(* IEC 61131-3 sources: plc-st-coding-agent/progress/evidence/f14_v11_public_20261113/jobs/custom_minimax-m27, 8 files *)

(* ---- public-easy-01.candidate_01.st ---- *)
(* ENGINEERING_CONTRACT
+--------------------------------------------------------------------------------------+
| Output             | Activation                | Retention | Reset/Deactivation    | Units |
|--------------------|---------------------------|-----------|-----------------------|-------|
| Pump_Motor         | bottleSensor in IDLE      | Hold      | cleaningConfirmButton | BOOL  |
| Filling_Valve      | cleaningConfirmButton     | Hold      | fillingConfirmButton  | BOOL  |
| Capping_Machine    | fillingConfirmButton      | Hold      | cappingConfirmButton  | BOOL  |
| Packing_Machine    | cappingConfirmButton      | Hold      | packingConfirmButton  | BOOL  |
| Completion_Light   | packingConfirmButton      | Hold      | finishedButton        | BOOL  |
+--------------------------------------------------------------------------------------+
| State Machine: IDLE->CLEANING->FILLING->CAPPING->PACKING->COMPLETED->IDLE           |
| All confirm inputs use R_TRIG for edge detection (same-scan priority preserved).     |
| Outputs are combinational to their active state; no edge memory needed.              |
| finishedButton only resets from COMPLETED state (PUB008).                            |
+--------------------------------------------------------------------------------------+
*)
(* CONTRACT_RULES [{"kind":"hold_until_reset","output":"Completion_Light","set_input":"packingConfirmButton","reset_input":"finishedButton"}] *)
FUNCTION_BLOCK BottleFillingLine
VAR_INPUT
    bottleSensor          : BOOL;
    cleaningConfirmButton : BOOL;
    fillingConfirmButton  : BOOL;
    cappingConfirmButton  : BOOL;
    packingConfirmButton  : BOOL;
    finishedButton        : BOOL;
END_VAR
VAR_OUTPUT
    Pump_Motor      : BOOL;
    Filling_Valve   : BOOL;
    Capping_Machine : BOOL;
    Packing_Machine : BOOL;
    Completion_Light: BOOL;
END_VAR
VAR
    eState : INT;
    IDLE      : INT := 0;
    CLEANING  : INT := 1;
    FILLING   : INT := 2;
    CAPPING   : INT := 3;
    PACKING   : INT := 4;
    COMPLETED : INT := 5;

    trigBottle   : R_TRIG;
    trigClean    : R_TRIG;
    trigFill     : R_TRIG;
    trigCap      : R_TRIG;
    trigPack     : R_TRIG;
    trigFinished : R_TRIG;
END_VAR

// Detect rising edges for all button inputs
trigBottle(CLK := bottleSensor);
trigClean(CLK := cleaningConfirmButton);
trigFill(CLK := fillingConfirmButton);
trigCap(CLK := cappingConfirmButton);
trigPack(CLK := packingConfirmButton);
trigFinished(CLK := finishedButton);

// State machine transitions
CASE eState OF
    IDLE:
        IF trigBottle.Q THEN
            eState := CLEANING;
        END_IF;

    CLEANING:
        IF trigClean.Q THEN
            eState := FILLING;
        END_IF;

    FILLING:
        IF trigFill.Q THEN
            eState := CAPPING;
        END_IF;

    CAPPING:
        IF trigCap.Q THEN
            eState := PACKING;
        END_IF;

    PACKING:
        IF trigPack.Q THEN
            eState := COMPLETED;
        END_IF;

    COMPLETED:
        IF trigFinished.Q THEN
            eState := IDLE;
        END_IF;
END_CASE;

// Output control based on current state
Pump_Motor       := (eState = CLEANING);
Filling_Valve    := (eState = FILLING);
Capping_Machine  := (eState = CAPPING);
Packing_Machine  := (eState = PACKING);
Completion_Light := (eState = COMPLETED);

END_FUNCTION_BLOCK

(* ---- public-easy-01.candidate_02.st ---- *)
(* ENGINEERING_CONTRACT
+--------------------------------------------------------------------------------------+
| Output             | Activation                | Retention | Reset/Deactivation    | Units |
|--------------------|---------------------------|-----------|-----------------------|-------|
| Pump_Motor         | bottleSensor in IDLE      | Hold      | cleaningConfirmButton | BOOL  |
| Filling_Valve      | cleaningConfirmButton     | Hold      | fillingConfirmButton  | BOOL  |
| Capping_Machine    | fillingConfirmButton      | Hold      | cappingConfirmButton  | BOOL  |
| Packing_Machine    | cappingConfirmButton      | Hold      | packingConfirmButton  | BOOL  |
| Completion_Light   | packingConfirmButton      | Hold      | finishedButton        | BOOL  |
+--------------------------------------------------------------------------------------+
| State Machine: IDLE->CLEANING->FILLING->CAPPING->PACKING->COMPLETED->IDLE           |
| All confirm inputs use R_TRIG for edge detection (same-scan priority preserved).     |
| Outputs are combinational to their active state; no edge memory needed.              |
| finishedButton only resets from COMPLETED state (PUB008).                            |
+--------------------------------------------------------------------------------------+
*)
(* CONTRACT_RULES [{"kind":"hold_until_reset","output":"Completion_Light","set_input":"packingConfirmButton","reset_input":"finishedButton"}] *)
FUNCTION_BLOCK BottleFillingLine
VAR_INPUT
    bottleSensor          : BOOL;
    cleaningConfirmButton : BOOL;
    fillingConfirmButton  : BOOL;
    cappingConfirmButton  : BOOL;
    packingConfirmButton  : BOOL;
    finishedButton        : BOOL;
END_VAR
VAR_OUTPUT
    Pump_Motor      : BOOL;
    Filling_Valve   : BOOL;
    Capping_Machine : BOOL;
    Packing_Machine : BOOL;
    Completion_Light: BOOL;
END_VAR
VAR
    eState : INT;

    trigBottle   : R_TRIG;
    trigClean    : R_TRIG;
    trigFill     : R_TRIG;
    trigCap      : R_TRIG;
    trigPack     : R_TRIG;
    trigFinished : R_TRIG;
END_VAR
VAR CONSTANT
    IDLE      : INT := 0;
    CLEANING  : INT := 1;
    FILLING   : INT := 2;
    CAPPING   : INT := 3;
    PACKING   : INT := 4;
    COMPLETED : INT := 5;
END_VAR

// Detect rising edges for all button inputs
trigBottle(CLK := bottleSensor);
trigClean(CLK := cleaningConfirmButton);
trigFill(CLK := fillingConfirmButton);
trigCap(CLK := cappingConfirmButton);
trigPack(CLK := packingConfirmButton);
trigFinished(CLK := finishedButton);

// State machine transitions
CASE eState OF
    IDLE:
        IF trigBottle.Q THEN
            eState := CLEANING;
        END_IF;

    CLEANING:
        IF trigClean.Q THEN
            eState := FILLING;
        END_IF;

    FILLING:
        IF trigFill.Q THEN
            eState := CAPPING;
        END_IF;

    CAPPING:
        IF trigCap.Q THEN
            eState := PACKING;
        END_IF;

    PACKING:
        IF trigPack.Q THEN
            eState := COMPLETED;
        END_IF;

    COMPLETED:
        IF trigFinished.Q THEN
            eState := IDLE;
        END_IF;
END_CASE;

// Output control based on current state
Pump_Motor       := (eState = CLEANING);
Filling_Valve    := (eState = FILLING);
Capping_Machine  := (eState = CAPPING);
Packing_Machine  := (eState = PACKING);
Completion_Light := (eState = COMPLETED);

END_FUNCTION_BLOCK

(* ---- public-easy-01.raw_candidate_01.st ---- *)
(* ENGINEERING_CONTRACT
+--------------------------------------------------------------------------------------+
| Output             | Activation                | Retention | Reset/Deactivation    | Units |
|--------------------|---------------------------|-----------|-----------------------|-------|
| Pump_Motor         | bottleSensor in IDLE      | Hold      | cleaningConfirmButton | BOOL  |
| Filling_Valve      | cleaningConfirmButton     | Hold      | fillingConfirmButton  | BOOL  |
| Capping_Machine    | fillingConfirmButton      | Hold      | cappingConfirmButton  | BOOL  |
| Packing_Machine    | cappingConfirmButton      | Hold      | packingConfirmButton  | BOOL  |
| Completion_Light   | packingConfirmButton      | Hold      | finishedButton        | BOOL  |
+--------------------------------------------------------------------------------------+
| State Machine: IDLE->CLEANING->FILLING->CAPPING->PACKING->COMPLETED->IDLE           |
| All confirm inputs use R_TRIG for edge detection (same-scan priority preserved).     |
| Outputs are combinational to their active state; no edge memory needed.              |
| finishedButton only resets from COMPLETED state (PUB008).                            |
+--------------------------------------------------------------------------------------+
*)
(* CONTRACT_RULES [{"kind":"hold_until_reset","output":"Completion_Light","set_input":"packingConfirmButton","reset_input":"finishedButton"}] *)
FUNCTION_BLOCK BottleFillingLine
VAR_INPUT
    bottleSensor          : BOOL;
    cleaningConfirmButton : BOOL;
    fillingConfirmButton  : BOOL;
    cappingConfirmButton  : BOOL;
    packingConfirmButton  : BOOL;
    finishedButton        : BOOL;
END_VAR
VAR_OUTPUT
    Pump_Motor      : BOOL;
    Filling_Valve   : BOOL;
    Capping_Machine : BOOL;
    Packing_Machine : BOOL;
    Completion_Light: BOOL;
END_VAR
VAR
    eState : INT;
    IDLE      : INT := 0;
    CLEANING  : INT := 1;
    FILLING   : INT := 2;
    CAPPING   : INT := 3;
    PACKING   : INT := 4;
    COMPLETED : INT := 5;

    trigBottle   : R_TRIG;
    trigClean    : R_TRIG;
    trigFill     : R_TRIG;
    trigCap      : R_TRIG;
    trigPack     : R_TRIG;
    trigFinished : R_TRIG;
END_VAR

// Detect rising edges for all button inputs
trigBottle(CLK := bottleSensor);
trigClean(CLK := cleaningConfirmButton);
trigFill(CLK := fillingConfirmButton);
trigCap(CLK := cappingConfirmButton);
trigPack(CLK := packingConfirmButton);
trigFinished(CLK := finishedButton);

// State machine transitions
CASE eState OF
    IDLE:
        IF trigBottle.Q THEN
            eState := CLEANING;
        END_IF;

    CLEANING:
        IF trigClean.Q THEN
            eState := FILLING;
        END_IF;

    FILLING:
        IF trigFill.Q THEN
            eState := CAPPING;
        END_IF;

    CAPPING:
        IF trigCap.Q THEN
            eState := PACKING;
        END_IF;

    PACKING:
        IF trigPack.Q THEN
            eState := COMPLETED;
        END_IF;

    COMPLETED:
        IF trigFinished.Q THEN
            eState := IDLE;
        END_IF;
END_CASE;

// Output control based on current state
Pump_Motor       := (eState = CLEANING);
Filling_Valve    := (eState = FILLING);
Capping_Machine  := (eState = CAPPING);
Packing_Machine  := (eState = PACKING);
Completion_Light := (eState = COMPLETED);

END_FUNCTION_BLOCK

(* ---- public-easy-01.raw_candidate_02.st ---- *)
(* ENGINEERING_CONTRACT
+--------------------------------------------------------------------------------------+
| Output             | Activation                | Retention | Reset/Deactivation    | Units |
|--------------------|---------------------------|-----------|-----------------------|-------|
| Pump_Motor         | bottleSensor in IDLE      | Hold      | cleaningConfirmButton | BOOL  |
| Filling_Valve      | cleaningConfirmButton     | Hold      | fillingConfirmButton  | BOOL  |
| Capping_Machine    | fillingConfirmButton      | Hold      | cappingConfirmButton  | BOOL  |
| Packing_Machine    | cappingConfirmButton      | Hold      | packingConfirmButton  | BOOL  |
| Completion_Light   | packingConfirmButton      | Hold      | finishedButton        | BOOL  |
+--------------------------------------------------------------------------------------+
| State Machine: IDLE->CLEANING->FILLING->CAPPING->PACKING->COMPLETED->IDLE           |
| All confirm inputs use R_TRIG for edge detection (same-scan priority preserved).     |
| Outputs are combinational to their active state; no edge memory needed.              |
| finishedButton only resets from COMPLETED state (PUB008).                            |
+--------------------------------------------------------------------------------------+
*)
(* CONTRACT_RULES [{"kind":"hold_until_reset","output":"Completion_Light","set_input":"packingConfirmButton","reset_input":"finishedButton"}] *)
FUNCTION_BLOCK BottleFillingLine
VAR_INPUT
    bottleSensor          : BOOL;
    cleaningConfirmButton : BOOL;
    fillingConfirmButton  : BOOL;
    cappingConfirmButton  : BOOL;
    packingConfirmButton  : BOOL;
    finishedButton        : BOOL;
END_VAR
VAR_OUTPUT
    Pump_Motor      : BOOL;
    Filling_Valve   : BOOL;
    Capping_Machine : BOOL;
    Packing_Machine : BOOL;
    Completion_Light: BOOL;
END_VAR
VAR
    eState : INT;

    trigBottle   : R_TRIG;
    trigClean    : R_TRIG;
    trigFill     : R_TRIG;
    trigCap      : R_TRIG;
    trigPack     : R_TRIG;
    trigFinished : R_TRIG;
END_VAR
VAR CONSTANT
    IDLE      : INT := 0;
    CLEANING  : INT := 1;
    FILLING   : INT := 2;
    CAPPING   : INT := 3;
    PACKING   : INT := 4;
    COMPLETED : INT := 5;
END_VAR

// Detect rising edges for all button inputs
trigBottle(CLK := bottleSensor);
trigClean(CLK := cleaningConfirmButton);
trigFill(CLK := fillingConfirmButton);
trigCap(CLK := cappingConfirmButton);
trigPack(CLK := packingConfirmButton);
trigFinished(CLK := finishedButton);

// State machine transitions
CASE eState OF
    IDLE:
        IF trigBottle.Q THEN
            eState := CLEANING;
        END_IF;

    CLEANING:
        IF trigClean.Q THEN
            eState := FILLING;
        END_IF;

    FILLING:
        IF trigFill.Q THEN
            eState := CAPPING;
        END_IF;

    CAPPING:
        IF trigCap.Q THEN
            eState := PACKING;
        END_IF;

    PACKING:
        IF trigPack.Q THEN
            eState := COMPLETED;
        END_IF;

    COMPLETED:
        IF trigFinished.Q THEN
            eState := IDLE;
        END_IF;
END_CASE;

// Output control based on current state
Pump_Motor       := (eState = CLEANING);
Filling_Valve    := (eState = FILLING);
Capping_Machine  := (eState = CAPPING);
Packing_Machine  := (eState = PACKING);
Completion_Light := (eState = COMPLETED);

END_FUNCTION_BLOCK

(* ---- public-easy-02.candidate_01.st ---- *)
(* ENGINEERING_CONTRACT:
 * - Inputs: value (DWORD, 32-bit), sampled every scan cycle
 * - Rising edge: prev=0 AND current=1 → risingBits = value AND NOT prevValue
 * - Falling edge: prev=1 AND current=0 → fallingBits = NOT value AND prevValue
 * - hasChanged: retention until next scan, set when value <> prevValue
 * - hasRisingEdges: combinational, true when risingBits <> 0
 * - hasFallingEdges: combinational, true when fallingBits <> 0
 * - risingBits/fallingBits: stored per-bit edge indicators, latching across scans
 * - noOfRisingBits/noOfFallingBits: USINT count of set bits in edge bitmasks
 * - Units: bit positions 0-31, counts 0-32
 * - Initialization: prevValue defaults to 0; first scan treats 0→1 as rising edges
 * - No explicit reset; state evolves per scan with prevValue update
 * - PUB001: Input value, edge detection logic, output reporting
 *)

(* CONTRACT_RULES [] *)

FUNCTION_BLOCK FB_DualWordEdgeDetection
VAR_INPUT
    value : DWORD;
END_VAR

VAR_OUTPUT
    hasChanged      : BOOL;
    hasRisingEdges  : BOOL;
    risingBits      : DWORD;
    noOfRisingBits  : USINT;
    hasFallingEdges : BOOL;
    fallingBits     : DWORD;
    noOfFallingBits : USINT;
END_VAR

VAR
    prevValue : DWORD;
END_VAR

VAR_TEMP
    tmp_i     : USINT;
END_VAR

    // Detect rising edges: current=1 AND previous=0
    risingBits := value AND NOT prevValue;

    // Detect falling edges: previous=1 AND current=0
    fallingBits := NOT value AND prevValue;

    // Report change detection
    hasChanged := value <> prevValue;

    // Report edge occurrence flags
    hasRisingEdges := risingBits <> 0;
    hasFallingEdges := fallingBits <> 0;

    // Count rising bits (0-32)
    noOfRisingBits := 0;
    FOR tmp_i := 0 TO 31 DO
        IF (risingBits AND (1 SHL tmp_i)) <> 0 THEN
            noOfRisingBits := noOfRisingBits + 1;
        END_IF;
    END_FOR;

    // Count falling bits (0-32)
    noOfFallingBits := 0;
    FOR tmp_i := 0 TO 31 DO
        IF (fallingBits AND (1 SHL tmp_i)) <> 0 THEN
            noOfFallingBits := noOfFallingBits + 1;
        END_IF;
    END_FOR;

    // Store current value for next scan comparison
    prevValue := value;
END_FUNCTION_BLOCK

(* ---- public-easy-02.candidate_02.st ---- *)
(* ENGINEERING_CONTRACT:
 * - Inputs: value (DWORD, 32-bit), sampled every scan cycle
 * - Rising edge: prev=0 AND current=1 → risingBits = value AND NOT prevValue
 * - Falling edge: prev=1 AND current=0 → fallingBits = NOT value AND prevValue
 * - hasChanged: retention until next scan, set when value <> prevValue
 * - hasRisingEdges: combinational, true when risingBits <> 0
 * - hasFallingEdges: combinational, true when fallingBits <> 0
 * - risingBits/fallingBits: stored per-bit edge indicators, latching across scans
 * - noOfRisingBits/noOfFallingBits: USINT count of set bits in edge bitmasks
 * - Units: bit positions 0-31, counts 0-32
 * - Initialization: prevValue defaults to 0; first scan treats 0→1 as rising edges
 * - No explicit reset; state evolves per scan with prevValue update
 * - PUB001: Input value, edge detection logic, output reporting
 *)

(* CONTRACT_RULES [] *)

FUNCTION_BLOCK FB_DualWordEdgeDetection
VAR_INPUT
    value : DWORD;
END_VAR

VAR_OUTPUT
    hasChanged      : BOOL;
    hasRisingEdges  : BOOL;
    risingBits      : DWORD;
    noOfRisingBits  : USINT;
    hasFallingEdges : BOOL;
    fallingBits     : DWORD;
    noOfFallingBits : USINT;
END_VAR

VAR
    prevValue : DWORD;
END_VAR

VAR_TEMP
    tmp_i     : USINT;
END_VAR

    // Detect rising edges: current=1 AND previous=0
    risingBits := value AND NOT prevValue;

    // Detect falling edges: previous=1 AND current=0
    fallingBits := NOT value AND prevValue;

    // Report change detection
    hasChanged := value <> prevValue;

    // Report edge occurrence flags
    hasRisingEdges := risingBits <> 0;
    hasFallingEdges := fallingBits <> 0;

    // Count rising bits (0-32)
    noOfRisingBits := 0;
    FOR tmp_i := 0 TO 31 DO
        IF (risingBits AND SHL(1, tmp_i)) <> 0 THEN
            noOfRisingBits := noOfRisingBits + 1;
        END_IF;
    END_FOR;

    // Count falling bits (0-32)
    noOfFallingBits := 0;
    FOR tmp_i := 0 TO 31 DO
        IF (fallingBits AND SHL(1, tmp_i)) <> 0 THEN
            noOfFallingBits := noOfFallingBits + 1;
        END_IF;
    END_FOR;

    // Store current value for next scan comparison
    prevValue := value;
END_FUNCTION_BLOCK

(* ---- public-easy-02.raw_candidate_01.st ---- *)
(* ENGINEERING_CONTRACT:
 * - Inputs: value (DWORD, 32-bit), sampled every scan cycle
 * - Rising edge: prev=0 AND current=1 → risingBits = value AND NOT prevValue
 * - Falling edge: prev=1 AND current=0 → fallingBits = NOT value AND prevValue
 * - hasChanged: retention until next scan, set when value <> prevValue
 * - hasRisingEdges: combinational, true when risingBits <> 0
 * - hasFallingEdges: combinational, true when fallingBits <> 0
 * - risingBits/fallingBits: stored per-bit edge indicators, latching across scans
 * - noOfRisingBits/noOfFallingBits: USINT count of set bits in edge bitmasks
 * - Units: bit positions 0-31, counts 0-32
 * - Initialization: prevValue defaults to 0; first scan treats 0→1 as rising edges
 * - No explicit reset; state evolves per scan with prevValue update
 * - PUB001: Input value, edge detection logic, output reporting
 *)

(* CONTRACT_RULES [] *)

FUNCTION_BLOCK FB_DualWordEdgeDetection
VAR_INPUT
    value : DWORD;
END_VAR

VAR_OUTPUT
    hasChanged      : BOOL;
    hasRisingEdges  : BOOL;
    risingBits      : DWORD;
    noOfRisingBits  : USINT;
    hasFallingEdges : BOOL;
    fallingBits     : DWORD;
    noOfFallingBits : USINT;
END_VAR

VAR
    prevValue : DWORD;
END_VAR

VAR_TEMP
    tmp_i     : USINT;
END_VAR

    // Detect rising edges: current=1 AND previous=0
    risingBits := value AND NOT prevValue;

    // Detect falling edges: previous=1 AND current=0
    fallingBits := NOT value AND prevValue;

    // Report change detection
    hasChanged := value <> prevValue;

    // Report edge occurrence flags
    hasRisingEdges := risingBits <> 0;
    hasFallingEdges := fallingBits <> 0;

    // Count rising bits (0-32)
    noOfRisingBits := 0;
    FOR tmp_i := 0 TO 31 DO
        IF (risingBits AND (1 SHL tmp_i)) <> 0 THEN
            noOfRisingBits := noOfRisingBits + 1;
        END_IF;
    END_FOR;

    // Count falling bits (0-32)
    noOfFallingBits := 0;
    FOR tmp_i := 0 TO 31 DO
        IF (fallingBits AND (1 SHL tmp_i)) <> 0 THEN
            noOfFallingBits := noOfFallingBits + 1;
        END_IF;
    END_FOR;

    // Store current value for next scan comparison
    prevValue := value;
END_FUNCTION_BLOCK

(* ---- public-easy-02.raw_candidate_02.st ---- *)
(* ENGINEERING_CONTRACT:
 * - Inputs: value (DWORD, 32-bit), sampled every scan cycle
 * - Rising edge: prev=0 AND current=1 → risingBits = value AND NOT prevValue
 * - Falling edge: prev=1 AND current=0 → fallingBits = NOT value AND prevValue
 * - hasChanged: retention until next scan, set when value <> prevValue
 * - hasRisingEdges: combinational, true when risingBits <> 0
 * - hasFallingEdges: combinational, true when fallingBits <> 0
 * - risingBits/fallingBits: stored per-bit edge indicators, latching across scans
 * - noOfRisingBits/noOfFallingBits: USINT count of set bits in edge bitmasks
 * - Units: bit positions 0-31, counts 0-32
 * - Initialization: prevValue defaults to 0; first scan treats 0→1 as rising edges
 * - No explicit reset; state evolves per scan with prevValue update
 * - PUB001: Input value, edge detection logic, output reporting
 *)

(* CONTRACT_RULES [] *)

FUNCTION_BLOCK FB_DualWordEdgeDetection
VAR_INPUT
    value : DWORD;
END_VAR

VAR_OUTPUT
    hasChanged      : BOOL;
    hasRisingEdges  : BOOL;
    risingBits      : DWORD;
    noOfRisingBits  : USINT;
    hasFallingEdges : BOOL;
    fallingBits     : DWORD;
    noOfFallingBits : USINT;
END_VAR

VAR
    prevValue : DWORD;
END_VAR

VAR_TEMP
    tmp_i     : USINT;
END_VAR

    // Detect rising edges: current=1 AND previous=0
    risingBits := value AND NOT prevValue;

    // Detect falling edges: previous=1 AND current=0
    fallingBits := NOT value AND prevValue;

    // Report change detection
    hasChanged := value <> prevValue;

    // Report edge occurrence flags
    hasRisingEdges := risingBits <> 0;
    hasFallingEdges := fallingBits <> 0;

    // Count rising bits (0-32)
    noOfRisingBits := 0;
    FOR tmp_i := 0 TO 31 DO
        IF (risingBits AND SHL(1, tmp_i)) <> 0 THEN
            noOfRisingBits := noOfRisingBits + 1;
        END_IF;
    END_FOR;

    // Count falling bits (0-32)
    noOfFallingBits := 0;
    FOR tmp_i := 0 TO 31 DO
        IF (fallingBits AND SHL(1, tmp_i)) <> 0 THEN
            noOfFallingBits := noOfFallingBits + 1;
        END_IF;
    END_FOR;

    // Store current value for next scan comparison
    prevValue := value;
END_FUNCTION_BLOCK
